Fanuc KAREL source: KO00133.KL

PROGRAM KO00133
%NOLOCKGROUP
VAR
  R: REAL
  CFG: CONFIG
  OUT: XYZWPR
  N: INTEGER
BEGIN
  N = 1
  R = 2.0
  CFG.CFG_FLIP = TRUE
  OUT = POS(R, N, R, R, R, R, CFG)
END KO00133
